(* IEC 61131-3 sources: PLC-ST-Learning/examples/datacenter_control_expert, 5 files *)

(* ---- 01_Types.st ---- *)
(* IEC reference declarations. Create these DDTs in Control Expert's Data Editor.
   This file is NOT an XDB/XEF import file. Indices are always 1..16. *)
TYPE T_DC_TrainStatus :
STRUCT
    Available : BOOL;
    Ready : BOOL;
    Loaded : BOOL;
    ChillerRunning : BOOL;
    Starting : BOOL;
    Stopping : BOOL;
    CanStop : BOOL;
    Fault : BOOL;
    State : INT;
    FaultCode : INT;
END_STRUCT
END_TYPE

TYPE T_DC_StatusArray : ARRAY [1..16] OF T_DC_TrainStatus; END_TYPE
TYPE T_DC_BoolArray : ARRAY [1..16] OF BOOL; END_TYPE
TYPE T_DC_HoursArray : ARRAY [1..16] OF REAL; END_TYPE

TYPE T_DC_TrainIO :
STRUCT
    RemoteAuto : BOOL;
    Maintenance : BOOL;
    RunPermit : BOOL;
    PowerAvailable : BOOL;
    HardTrip : BOOL;
    ChillerFault : BOOL;
    WaterEquipmentFault : BOOL;
    ValveOpenFb : BOOL;
    ValveClosedFb : BOOL;
    ChwPumpRunFb : BOOL;
    CwPumpRunFb : BOOL;
    ChwFlowOk : BOOL;
    CwFlowOk : BOOL;
    TowerReadyFb : BOOL;
    ChillerRunFb : BOOL;
    LoadedFb : BOOL;
    LoadPermit : BOOL;
    Reset : BOOL;
    OpenValvesCmd : BOOL;
    RunChwPumpCmd : BOOL;
    RunCwPumpCmd : BOOL;
    RequestTowerCmd : BOOL;
    RunChillerCmd : BOOL;
    EnableLoadCmd : BOOL;
END_STRUCT
END_TYPE
TYPE T_DC_IOArray : ARRAY [1..16] OF T_DC_TrainIO; END_TYPE

(* ---- 02_FB_DC_Train.st ---- *)
(* Reference DFB: dedicated water equipment per chiller.
   Split declarations and body into a Control Expert DFB; see the Chinese guide.
   All commands are level signals; adapt to vendor start/stop interfaces separately. *)
FUNCTION_BLOCK FB_DC_Train
VAR_INPUT
    FirstScan : BOOL;
    RequestRun : BOOL;
    Reset : BOOL;
    RemoteAuto : BOOL;
    Maintenance : BOOL;
    RunPermit : BOOL;
    PowerAvailable : BOOL; (* Real per-train power feedback, distinct from process trips *)
    HardTrip : BOOL;
    ChillerFault : BOOL;
    WaterEquipmentFault : BOOL;
    ValveOpenFb : BOOL; (* Combined chilled/condenser valve open proof *)
    ValveClosedFb : BOOL;
    ChwPumpRunFb : BOOL;
    CwPumpRunFb : BOOL;
    ChwFlowOk : BOOL;
    CwFlowOk : BOOL;
    TowerReadyFb : BOOL; (* From tower controller; includes local fan staging *)
    ChillerRunFb : BOOL;
    LoadedFb : BOOL; (* Must be real ready/capacity feedback, not command echo *)
    LoadPermit : BOOL;
    MinOff : TIME := T#10m;
    MinOn : TIME := T#10m;
    ValveTimeout : TIME := T#60s;
    PumpTimeout : TIME := T#30s;
    FlowStable : TIME := T#15s;
    FlowTimeout : TIME := T#90s;
    FlowLossDelay : TIME := T#2s;
    CapacityLossDelay : TIME := T#10s;
    TowerTimeout : TIME := T#120s;
    ChillerTimeout : TIME := T#180s;
    LoadTimeout : TIME := T#180s;
    UnloadTimeout : TIME := T#120s;
    StopTimeout : TIME := T#180s;
    PostRun : TIME := T#180s;
END_VAR
VAR_OUTPUT
    OpenValves : BOOL;
    RunChwPump : BOOL;
    RunCwPump : BOOL;
    RequestTower : BOOL;
    RunChiller : BOOL;
    EnableLoad : BOOL;
    Status : T_DC_TrainStatus;
    UnloadTimedOut : BOOL;
    StopTimedOut : BOOL;
END_VAR
VAR
    State : INT;
    FaultLatched : BOOL;
    FaultCode : INT;
    OldReset : BOOL;
    ResetEdge : BOOL;
    WaterOk : BOOL;
    ConfigOk : BOOL;
    ControlledTrip : BOOL;
    tmOff : TON;
    tmOn : TON;
    tmValveOpen : TON;
    tmPump : TON;
    tmFlowStable : TON;
    tmFlowWait : TON;
    tmFlowLoss : TON;
    tmCapacityLoss : TON;
    tmTower : TON;
    tmChiller : TON;
    tmLoad : TON;
    tmUnload : TON;
    tmStop : TON;
    tmPost : TON;
    tmPumpStop : TON;
    tmValveClose : TON;
END_VAR

ResetEdge := Reset AND NOT OldReset;
OldReset := Reset;
ConfigOk := (MinOff > T#0s) AND (MinOn > T#0s)
    AND (ValveTimeout > T#0s) AND (PumpTimeout > T#0s)
    AND (FlowStable > T#0s) AND (FlowTimeout > FlowStable)
    AND (FlowLossDelay >= T#0s) AND (CapacityLossDelay > T#0s)
    AND (TowerTimeout > T#0s)
    AND (ChillerTimeout > T#0s) AND (LoadTimeout > T#0s)
    AND (UnloadTimeout > T#0s) AND (StopTimeout > T#0s)
    AND (PostRun > T#0s);
WaterOk := ValveOpenFb AND ChwPumpRunFb AND CwPumpRunFb
    AND ChwFlowOk AND CwFlowOk;

(* Non-retained state is reconstructed from real feedback, never retained commands. *)
IF FirstScan THEN
    OldReset := Reset;
    ResetEdge := FALSE;
    State := 0;
    FaultLatched := FALSE;
    FaultCode := 0;
    UnloadTimedOut := FALSE;
    StopTimedOut := FALSE;
    IF ChillerRunFb THEN
        IF LoadedFb THEN State := 70; ELSE State := 60; END_IF;
    ELSIF ChwPumpRunFb OR CwPumpRunFb THEN
        State := 100;
    ELSIF ValveOpenFb THEN
        State := 120;
    END_IF;
END_IF;

(* Call EVERY timer exactly once per scan, even while idle or faulted. *)
tmOff(IN := NOT ChillerRunFb AND NOT FirstScan, PT := MinOff);
tmOn(IN := ChillerRunFb AND NOT FirstScan, PT := MinOn);
tmValveOpen(IN := (State = 10) AND NOT FirstScan, PT := ValveTimeout);
tmPump(IN := (State = 20) AND NOT FirstScan, PT := PumpTimeout);
tmFlowStable(IN := WaterOk AND NOT FirstScan, PT := FlowStable);
tmFlowWait(IN := (State = 30) AND NOT FirstScan, PT := FlowTimeout);
tmFlowLoss(IN := (State >= 50) AND (State <= 80) AND NOT WaterOk
    AND NOT FirstScan, PT := FlowLossDelay);
tmCapacityLoss(IN := (State = 70) AND NOT LoadedFb AND NOT FirstScan,
    PT := CapacityLossDelay);
tmTower(IN := (State = 40) AND NOT FirstScan, PT := TowerTimeout);
tmChiller(IN := (State = 50) AND NOT FirstScan, PT := ChillerTimeout);
tmLoad(IN := (State = 60) AND NOT FirstScan, PT := LoadTimeout);
tmUnload(IN := (State = 80) AND NOT FirstScan, PT := UnloadTimeout);
tmStop(IN := (State = 90) AND NOT FirstScan, PT := StopTimeout);
tmPost(IN := (State = 100) AND NOT FirstScan, PT := PostRun);
tmPumpStop(IN := (State = 110) AND NOT FirstScan, PT := PumpTimeout);
tmValveClose(IN := (State = 120) AND NOT FirstScan, PT := ValveTimeout);

IF ResetEdge AND NOT ChillerRunFb AND NOT ChwPumpRunFb AND NOT CwPumpRunFb
    AND ValveClosedFb AND NOT ValveOpenFb AND NOT LoadedFb
    AND NOT ChillerFault AND NOT WaterEquipmentFault AND RunPermit
    AND NOT HardTrip AND RemoteAuto AND PowerAvailable AND ConfigOk
    AND ((State = 0) OR (State = 900)) THEN
    FaultLatched := FALSE;
    FaultCode := 0;
    UnloadTimedOut := FALSE;
    StopTimedOut := FALSE;
    State := 0;
END_IF;

ControlledTrip := FALSE;
IF NOT ConfigOk THEN FaultCode := 1; ControlledTrip := TRUE;
ELSIF NOT RunPermit AND (((State > 0) AND (State < 90)) OR ChillerRunFb) THEN
    FaultCode := 2; ControlledTrip := TRUE;
ELSIF ChillerFault THEN FaultCode := 3; ControlledTrip := TRUE;
ELSIF WaterEquipmentFault THEN FaultCode := 4; ControlledTrip := TRUE;
ELSIF (State >= 50) AND (State <= 80) AND NOT ValveOpenFb THEN
    FaultCode := 5; ControlledTrip := TRUE;
ELSIF tmFlowLoss.Q THEN FaultCode := 6; ControlledTrip := TRUE;
ELSIF (State >= 50) AND (State <= 80) AND NOT TowerReadyFb THEN
    FaultCode := 7; ControlledTrip := TRUE;
ELSIF ((State = 60) OR (State = 70) OR (State = 80)) AND NOT ChillerRunFb THEN
    FaultCode := 8; ControlledTrip := TRUE;
ELSIF tmCapacityLoss.Q THEN
    FaultCode := 9; ControlledTrip := TRUE;
ELSIF LoadedFb AND NOT ChillerRunFb THEN
    FaultCode := 10; ControlledTrip := TRUE;
ELSIF ValveOpenFb AND ValveClosedFb THEN
    FaultCode := 11; ControlledTrip := TRUE;
ELSIF ChillerRunFb AND ((State < 50) OR ((State >= 100) AND (State <= 120))
    OR (State = 900)) THEN
    FaultCode := 14; ControlledTrip := TRUE;
END_IF;

(* Hardwired safeties remain independent. A hard trip removes ALL commands. *)
IF HardTrip THEN
    FaultLatched := TRUE;
    FaultCode := 12;
    State := 900;
ELSIF NOT RemoteAuto THEN
    IF ChillerRunFb OR ChwPumpRunFb OR CwPumpRunFb
        OR ((State > 0) AND (State < 900)) THEN
        FaultLatched := TRUE; FaultCode := 13;
    END_IF;
    IF FaultLatched THEN State := 900; ELSE State := 0; END_IF;
ELSIF NOT PowerAvailable THEN
    (* Expected loss of supply is not a device-fault latch. Existing faults persist. *)
    State := 910;
ELSIF ControlledTrip THEN
    FaultLatched := TRUE;
    IF ChillerRunFb AND (State >= 100) THEN
        State := 90;
    ELSIF (State < 90) OR (State = 900) THEN
        IF ChillerRunFb THEN State := 90;
        ELSIF ChwPumpRunFb OR CwPumpRunFb THEN State := 100;
        ELSIF NOT ValveClosedFb THEN State := 120;
        ELSE State := 900;
        END_IF;
    END_IF;
END_IF;

(* Normal request withdrawal honors MinOn. Startup cancellation needs no MinOn. *)
IF NOT FirstScan AND NOT RequestRun AND NOT ControlledTrip AND NOT HardTrip
    AND RemoteAuto AND PowerAvailable AND (State > 0) AND (State < 80) THEN
    IF (State = 70) AND tmOn.Q THEN State := 80;
    ELSIF State = 10 THEN State := 120;
    ELSIF (State >= 20) AND (State <= 40) THEN State := 100;
    ELSIF (State = 50) OR (State = 60) THEN
        IF ChillerRunFb THEN State := 80; ELSE State := 100; END_IF;
    END_IF;
END_IF;

IF NOT HardTrip AND RemoteAuto AND PowerAvailable THEN
    CASE State OF
    0:
        IF ChillerRunFb OR ChwPumpRunFb OR CwPumpRunFb OR LoadedFb THEN
            FaultLatched := TRUE; FaultCode := 14;
            IF ChillerRunFb THEN State := 90; ELSE State := 100; END_IF;
        ELSIF RequestRun AND NOT FaultLatched AND NOT Maintenance
            AND RunPermit AND ConfigOk AND tmOff.Q AND ValveClosedFb THEN
            State := 10;
        END_IF;
    10:
        IF ValveOpenFb AND NOT ValveClosedFb THEN State := 20;
        ELSIF tmValveOpen.Q THEN FaultLatched := TRUE; FaultCode := 20; State := 120;
        END_IF;
    20:
        IF ChwPumpRunFb AND CwPumpRunFb THEN State := 30;
        ELSIF tmPump.Q THEN FaultLatched := TRUE; FaultCode := 21; State := 100;
        END_IF;
    30:
        IF tmFlowStable.Q THEN State := 40;
        ELSIF tmFlowWait.Q THEN FaultLatched := TRUE; FaultCode := 22; State := 100;
        END_IF;
    40:
        IF TowerReadyFb AND tmFlowStable.Q THEN State := 50;
        ELSIF tmTower.Q THEN FaultLatched := TRUE; FaultCode := 23; State := 100;
        END_IF;
    50:
        IF ChillerRunFb THEN State := 60;
        ELSIF tmChiller.Q THEN FaultLatched := TRUE; FaultCode := 24; State := 90;
        END_IF;
    60:
        IF LoadedFb AND LoadPermit AND tmFlowStable.Q THEN State := 70;
        ELSIF tmLoad.Q THEN FaultLatched := TRUE; FaultCode := 25; State := 80;
        END_IF;
    70:
        (* Loss of load permission unloads through the normal stop path. *)
        IF NOT LoadPermit THEN
            FaultLatched := TRUE; FaultCode := 26; State := 80;
        END_IF;
    80:
        IF NOT LoadedFb THEN State := 90;
        ELSIF tmUnload.Q THEN
            UnloadTimedOut := TRUE; FaultLatched := TRUE; FaultCode := 27; State := 90;
        END_IF;
    90:
        (* A stuck run feedback MUST NOT be treated as a stopped chiller. *)
        IF NOT ChillerRunFb THEN State := 100;
        ELSIF tmStop.Q THEN
            StopTimedOut := TRUE; FaultLatched := TRUE; FaultCode := 28;
        END_IF;
    100:
        IF ChillerRunFb THEN
            FaultLatched := TRUE; FaultCode := 29; State := 90;
        ELSIF tmPost.Q THEN State := 110;
        END_IF;
    110:
        IF NOT ChwPumpRunFb AND NOT CwPumpRunFb THEN State := 120;
        ELSIF tmPumpStop.Q THEN
            FaultLatched := TRUE; FaultCode := 30;
            (* Keep valves open until BOTH pumps really stop. *)
        END_IF;
    120:
        IF ChillerRunFb OR ChwPumpRunFb OR CwPumpRunFb THEN
            FaultLatched := TRUE; FaultCode := 31;
            IF ChillerRunFb THEN State := 90; ELSE State := 110; END_IF;
        ELSIF ValveClosedFb AND NOT ValveOpenFb THEN
            IF FaultLatched THEN State := 900; ELSE State := 0; END_IF;
        ELSIF tmValveClose.Q THEN
            FaultLatched := TRUE; FaultCode := 32;
        END_IF;
    900:
        (* No automatic reset/retry. A real reset edge at a safe rest is required. *)
        IF ChillerRunFb THEN State := 90;
        ELSIF ChwPumpRunFb OR CwPumpRunFb THEN State := 100;
        END_IF;
    910:
        (* Re-establish a safe rest before allowing the fleet to restart this train. *)
        IF ChillerRunFb THEN State := 90;
        ELSIF ChwPumpRunFb OR CwPumpRunFb THEN State := 100;
        ELSIF NOT ValveClosedFb THEN State := 120;
        ELSIF FaultLatched THEN State := 900;
        ELSE State := 0;
        END_IF;
    ELSE
        FaultLatched := TRUE; FaultCode := 99;
        IF ChillerRunFb THEN State := 90; ELSE State := 100; END_IF;
    END_CASE;
END_IF;

OpenValves := (State >= 10) AND (State <= 110);
RunChwPump := (State >= 20) AND (State <= 100);
RunCwPump := RunChwPump;
RequestTower := (State >= 40) AND (State <= 100);
RunChiller := (State >= 50) AND (State <= 80);
EnableLoad := (((State = 60) AND tmFlowStable.Q) OR ((State = 70) AND WaterOk))
    AND LoadPermit AND TowerReadyFb AND ChillerRunFb AND NOT FaultLatched;
(* Physical interlocks cut chiller/load immediately; water may continue for post-run. *)
RunChiller := RunChiller AND RunPermit AND NOT ChillerFault
    AND NOT WaterEquipmentFault AND ValveOpenFb AND NOT tmFlowLoss.Q
    AND TowerReadyFb AND ConfigOk AND ((State <> 50) OR WaterOk);
IF HardTrip OR NOT RemoteAuto OR NOT PowerAvailable THEN
    OpenValves := FALSE; RunChwPump := FALSE; RunCwPump := FALSE;
    RequestTower := FALSE; RunChiller := FALSE; EnableLoad := FALSE;
END_IF;
EnableLoad := EnableLoad AND RunChiller;
Status.Available := RemoteAuto AND NOT Maintenance AND RunPermit
    AND PowerAvailable
    AND NOT HardTrip AND NOT ChillerFault AND NOT WaterEquipmentFault
    AND NOT FaultLatched AND ConfigOk;
Status.Ready := Status.Available AND (State = 0) AND tmOff.Q
    AND ValveClosedFb AND NOT ValveOpenFb AND NOT ChillerRunFb
    AND NOT ChwPumpRunFb AND NOT CwPumpRunFb AND NOT LoadedFb;
Status.Loaded := (State = 70) AND LoadedFb AND ChillerRunFb AND WaterOk
    AND TowerReadyFb AND LoadPermit AND NOT FaultLatched
    AND RemoteAuto AND RunPermit AND NOT HardTrip;
Status.ChillerRunning := ChillerRunFb;
Status.Starting := (State >= 10) AND (State <= 60);
Status.Stopping := (State >= 80) AND (State <= 120);
Status.CanStop := (State = 70) AND tmOn.Q;
Status.Fault := FaultLatched;
Status.State := State;
Status.FaultCode := FaultCode;
END_FUNCTION_BLOCK

(* ---- 03_FB_DC_Plant.st ---- *)
(* Fleet dispatch. Equal-capacity chillers; maximum 16.
   Call all Train DFBs BEFORE this DFB; requests take effect next PLC scan. *)
FUNCTION_BLOCK FB_DC_Plant
VAR_INPUT
    FirstScan : BOOL;
    Enable : BOOL;
    DisasterActive : BOOL; (* Recovery latch input, NOT a safety output *)
    InfrastructureReady : BOOL; (* Power, BMS authority, common water system ready *)
    AckRecovery : BOOL;
    AutoRecovery : BOOL := FALSE;
    ResetAlarm : BOOL;
    DemandValid : BOOL;
    Demand : INT; (* Desired duty count from BMS or validated demand regulator *)
    UnitCount : INT := 4;
    MaxDuty : INT := 3; (* N+1 reserve with four installed units *)
    MaxParallel : INT := 4; (* Electrical/hydraulic limit, includes rotation overlap *)
    RotateEnable : BOOL := TRUE;
    RotateNow : BOOL;
    Status : T_DC_StatusArray;
    RunHours : T_DC_HoursArray; (* External, validated RETAIN hour meters *)
    RecoveryStable : TIME := T#60s;
    StartSpacing : TIME := T#120s;
    DemandUpDelay : TIME := T#60s;
    DemandDownDelay : TIME := T#300s;
    RotationInterval : TIME := T#168h;
    RotationOverlap : TIME := T#60s;
    RotationTimeout : TIME := T#30m;
END_VAR
VAR_OUTPUT
    Request : T_DC_BoolArray;
    RecoveryHold : BOOL;
    Target : INT;
    RunningCount : INT;
    LoadedCount : INT;
    RequestedCount : INT;
    CapacityShortage : BOOL;
    NoStartCandidate : BOOL;
    ReserveUnavailable : BOOL;
    ConfigFault : BOOL;
    RotationBlocked : BOOL;
    RotationFailed : BOOL;
    RotationActive : BOOL;
    InvalidDemand : BOOL;
END_VAR
VAR
    i : INT;
    n : INT;
    Candidate : INT;
    StopCandidate : INT;
    RotOld : INT;
    RotNew : INT;
    RotPhase : INT; (* 0 idle; 1 start replacement; 2 old train shutting down *)
    ReadyCount : INT;
    OccupiedCount : INT;
    LastDemand : INT;
    RotationTarget : INT;
    Desired : INT;
    MinHours : REAL;
    MaxHours : REAL;
    Starting : BOOL;
    Stopping : BOOL;
    OldAck : BOOL;
    OldRotate : BOOL;
    OldReset : BOOL;
    AckEdge : BOOL;
    RotateEdge : BOOL;
    ResetEdge : BOOL;
    SpacingActive : BOOL;
    SpacingReset : BOOL;
    RotationClockReset : BOOL;
    ReplacementLoaded : BOOL;
    tmRecovery : TON;
    tmSpacing : TON;
    tmUp : TON;
    tmDown : TON;
    tmRotation : TON;
    tmOverlap : TON;
    tmRotationTimeout : TON;
END_VAR

ConfigFault := (UnitCount < 1) OR (UnitCount > 16) OR (MaxDuty < 1)
    OR (MaxDuty > UnitCount) OR (MaxParallel < MaxDuty)
    OR (MaxParallel > UnitCount) OR (RecoveryStable <= T#0s)
    OR (StartSpacing <= T#0s) OR (DemandUpDelay < T#0s)
    OR (DemandDownDelay < T#0s) OR (RotationInterval <= T#0s)
    OR (RotationOverlap <= T#0s) OR (RotationTimeout <= RotationOverlap);
n := UnitCount;
IF n < 1 THEN n := 1; END_IF;
IF n > 16 THEN n := 16; END_IF;
AckEdge := AckRecovery AND NOT OldAck;
RotateEdge := RotateNow AND NOT OldRotate;
ResetEdge := ResetAlarm AND NOT OldReset;
OldAck := AckRecovery; OldRotate := RotateNow; OldReset := ResetAlarm;

IF FirstScan THEN
    RecoveryHold := TRUE;
    Target := 0; LastDemand := -1;
    RotPhase := 0; RotOld := 0; RotNew := 0;
    SpacingActive := TRUE; SpacingReset := TRUE; RotationClockReset := TRUE;
    RotationFailed := FALSE;
    AckEdge := FALSE; RotateEdge := FALSE; ResetEdge := FALSE;
    (* Adopt operating trains; never replay a retained command array. *)
    FOR i := 1 TO 16 DO
        Request[i] := (i <= n) AND Status[i].Available
            AND (Status[i].ChillerRunning OR Status[i].Starting);
        IF Request[i] THEN Target := Target + 1; END_IF;
    END_FOR;
END_IF;
IF DisasterActive OR NOT InfrastructureReady THEN RecoveryHold := TRUE; END_IF;

(* Invalid demand freezes the current target; it MUST NOT become zero demand. *)
InvalidDemand := NOT DemandValid OR (Demand < 0) OR (Demand > MaxDuty);
Desired := Target;
IF NOT InvalidDemand THEN Desired := Demand; END_IF;
IF NOT Enable THEN Desired := 0; END_IF;

tmRecovery(IN := InfrastructureReady AND NOT DisasterActive AND NOT FirstScan,
    PT := RecoveryStable);
tmSpacing(IN := SpacingActive AND NOT SpacingReset AND NOT FirstScan, PT := StartSpacing);
tmUp(IN := Enable AND NOT InvalidDemand AND NOT RecoveryHold
    AND (Desired > Target) AND (Desired = LastDemand) AND NOT FirstScan,
    PT := DemandUpDelay);
tmDown(IN := NOT InvalidDemand AND NOT RecoveryHold AND (Desired < Target)
    AND (Desired = LastDemand) AND NOT FirstScan, PT := DemandDownDelay);
tmRotation(IN := Enable AND RotateEnable AND NOT RecoveryHold AND (Target > 0)
    AND (RotPhase = 0) AND NOT RotationClockReset AND NOT FirstScan,
    PT := RotationInterval);
ReplacementLoaded := FALSE;
IF (RotNew >= 1) AND (RotNew <= n) THEN
    ReplacementLoaded := Status[RotNew].Loaded;
END_IF;
tmOverlap(IN := (RotPhase = 1) AND ReplacementLoaded
    AND NOT FirstScan, PT := RotationOverlap);
tmRotationTimeout(IN := (RotPhase <> 0) AND NOT FirstScan, PT := RotationTimeout);
RotationClockReset := FALSE;
SpacingReset := FALSE;
IF tmSpacing.Q THEN SpacingActive := FALSE; END_IF;
IF ResetEdge THEN RotationFailed := FALSE; END_IF;
IF RecoveryHold AND tmRecovery.Q AND (AutoRecovery OR AckEdge) AND Enable
    AND NOT ConfigFault THEN
    RecoveryHold := FALSE;
    SpacingActive := TRUE;
    SpacingReset := TRUE;
END_IF;
IF NOT Enable THEN Target := 0;
ELSIF NOT RecoveryHold AND NOT ConfigFault THEN
    IF tmUp.Q OR tmDown.Q THEN Target := Desired; END_IF;
END_IF;
LastDemand := Desired;

RunningCount := 0; LoadedCount := 0; RequestedCount := 0;
ReadyCount := 0; OccupiedCount := 0;
Starting := FALSE; Stopping := FALSE;
FOR i := 1 TO 16 DO
    IF i <= n THEN
        IF Status[i].ChillerRunning THEN RunningCount := RunningCount + 1; END_IF;
        IF Status[i].Loaded THEN LoadedCount := LoadedCount + 1; END_IF;
        IF Status[i].Ready THEN ReadyCount := ReadyCount + 1; END_IF;
        IF NOT Status[i].Available THEN Request[i] := FALSE; END_IF;
        IF Request[i] THEN RequestedCount := RequestedCount + 1; END_IF;
        IF Request[i] OR Status[i].ChillerRunning OR Status[i].Starting THEN
            OccupiedCount := OccupiedCount + 1;
        END_IF;
        Starting := Starting OR Status[i].Starting;
        Stopping := Stopping OR Status[i].Stopping;
    ELSE
        Request[i] := FALSE;
    END_IF;
END_FOR;

(* Select least-hours available start and greatest-hours stoppable running train.
   Ascending index resolves ties deterministically. *)
Candidate := 0; StopCandidate := 0;
MinHours := 3.0E+38; MaxHours := -1.0;
FOR i := 1 TO n DO
    IF Status[i].Ready AND NOT Request[i] AND (RunHours[i] >= 0.0)
        AND (RunHours[i] < MinHours) THEN
        Candidate := i; MinHours := RunHours[i];
    END_IF;
    IF Request[i] AND Status[i].Loaded AND Status[i].CanStop
        AND (RunHours[i] >= 0.0) AND (RunHours[i] > MaxHours) THEN
        StopCandidate := i; MaxHours := RunHours[i];
    END_IF;
END_FOR;

RotationBlocked := FALSE;
IF RotPhase <> 0 THEN
    (* Bound indices before use. No reliance on short-circuit array evaluation. *)
    IF (RotOld < 1) OR (RotOld > n) OR (RotNew < 1) OR (RotNew > n) THEN
        RotPhase := 0; RotationFailed := TRUE; RotationClockReset := TRUE;
    ELSE
        IF ConfigFault OR RecoveryHold OR NOT Enable OR InvalidDemand
            OR (Target <> RotationTarget) THEN
            (* Keep the original running unit; cancel replacement normally. *)
            IF RotPhase = 1 THEN Request[RotNew] := FALSE; END_IF;
            RotPhase := 0; RotationClockReset := TRUE;
        ELSIF NOT Status[RotOld].Available THEN
            (* Original failed: replacement is now ordinary fault replacement. *)
            RotPhase := 0; RotationClockReset := TRUE;
        ELSIF NOT Status[RotNew].Available OR tmRotationTimeout.Q THEN
            IF RotPhase = 1 THEN Request[RotNew] := FALSE; END_IF;
            RotationFailed := TRUE; RotPhase := 0; RotationClockReset := TRUE;
        ELSIF RotPhase = 1 THEN
            IF Status[RotNew].Loaded AND tmOverlap.Q AND Status[RotOld].CanStop THEN
                Request[RotOld] := FALSE; RotPhase := 2;
            END_IF;
        ELSIF RotPhase = 2 THEN
            IF NOT Status[RotOld].ChillerRunning AND NOT Status[RotOld].Stopping THEN
                RotPhase := 0; RotationClockReset := TRUE;
            END_IF;
        END_IF;
    END_IF;
END_IF;

IF NOT ConfigFault AND NOT RecoveryHold AND Enable
    AND (RotPhase = 0) AND NOT Starting THEN
    IF RequestedCount < Target THEN
        (* Fault replacement bypasses demand debounce, not start spacing or MinOff.
           Failed trains may finish water post-run while a spare starts. *)
        IF (Candidate > 0) AND NOT SpacingActive AND (OccupiedCount < MaxParallel) THEN
            Request[Candidate] := TRUE;
            SpacingActive := TRUE;
            SpacingReset := TRUE;
        END_IF;
    ELSIF (RequestedCount > Target) AND NOT Stopping AND NOT InvalidDemand THEN
        IF StopCandidate > 0 THEN Request[StopCandidate] := FALSE; END_IF;
    ELSIF RotateEnable AND NOT InvalidDemand AND (RotateEdge OR tmRotation.Q) AND (Target > 0)
        AND (RequestedCount = Target) AND (LoadedCount >= Target)
        AND NOT Stopping THEN
        IF (Candidate > 0) AND (StopCandidate > 0) AND NOT SpacingActive
            AND (OccupiedCount < MaxParallel) THEN
            RotOld := StopCandidate; RotNew := Candidate; RotationTarget := Target;
            Request[RotNew] := TRUE; RotPhase := 1; SpacingActive := TRUE;
            SpacingReset := TRUE;
            RotationClockReset := TRUE;
        ELSE RotationBlocked := TRUE;
        END_IF;
    END_IF;
END_IF;
(* Disable is an orderly stop; hard stops are the individual Train.HardTrip input. *)
IF NOT Enable THEN
    FOR i := 1 TO 16 DO Request[i] := FALSE; END_FOR;
END_IF;

RotationActive := RotPhase <> 0;
RequestedCount := 0;
FOR i := 1 TO n DO
    IF Request[i] THEN RequestedCount := RequestedCount + 1; END_IF;
END_FOR;
CapacityShortage := Enable AND NOT InvalidDemand AND (LoadedCount < Demand);
NoStartCandidate := Enable AND NOT RecoveryHold
    AND (RequestedCount < Target) AND (Candidate = 0);
ReserveUnavailable := Enable AND (ReadyCount = 0);
END_FUNCTION_BLOCK

(* ---- 04_FB_DC_Demand.st ---- *)
(* Optional supervisory staging by chilled-water SUPPLY temperature.
   Native chiller controllers retain compressor/guide-vane/VFD modulation.
   Do not use with unequal-capacity units without a capacity-based redesign. *)
FUNCTION_BLOCK FB_DC_Demand
VAR_INPUT
    FirstScan : BOOL;
    Enable : BOOL;
    SensorValid : BOOL;
    SupplyTemperature : REAL;
    Setpoint : REAL := 7.0;
    AddBand : REAL := 0.7;
    ShedBand : REAL := 0.5;
    SensorMin : REAL := 0.0;
    SensorMax : REAL := 35.0;
    MinDuty : INT := 1;
    MaxDuty : INT := 3;
    LoadedCount : INT;
    PlantStable : BOOL; (* No starts, stops, rotation, or recovery in progress *)
    AddDelay : TIME := T#120s;
    ShedDelay : TIME := T#600s;
    SettleTime : TIME := T#600s;
END_VAR
VAR_OUTPUT
    Demand : INT;
    DemandValid : BOOL;
    SensorAlarm : BOOL;
    ConfigFault : BOOL;
END_VAR
VAR
    tmAdd : TON;
    tmShed : TON;
    tmSettle : TON;
    Settling : BOOL;
    ResetSettle : BOOL;
    CanAdjust : BOOL;
END_VAR

ConfigFault := (MinDuty < 0) OR (MaxDuty < 1) OR (MaxDuty > 16)
    OR (MinDuty > MaxDuty) OR (AddBand <= 0.0) OR (ShedBand <= 0.0)
    OR (SensorMin >= SensorMax) OR (Setpoint <= SensorMin)
    OR (Setpoint >= SensorMax) OR (AddDelay <= T#0s)
    OR (ShedDelay <= T#0s) OR (SettleTime <= T#0s);
(* Positive range tests also reject an IEEE NaN measurement. *)
SensorAlarm := NOT SensorValid OR NOT ((SupplyTemperature >= SensorMin)
    AND (SupplyTemperature <= SensorMax));
DemandValid := NOT ConfigFault AND NOT SensorAlarm;
IF FirstScan THEN
    Demand := MinDuty;
    IF (LoadedCount > MinDuty) AND (LoadedCount <= MaxDuty) THEN
        Demand := LoadedCount;
    END_IF;
    IF Demand < 0 THEN Demand := 0; END_IF;
    IF Demand > 16 THEN Demand := 16; END_IF;
    Settling := TRUE; ResetSettle := TRUE;
END_IF;
tmSettle(IN := Settling AND NOT ResetSettle AND NOT FirstScan, PT := SettleTime);
ResetSettle := FALSE;
IF tmSettle.Q THEN Settling := FALSE; END_IF;
CanAdjust := Enable AND DemandValid AND PlantStable AND NOT Settling
    AND (LoadedCount = Demand) AND NOT FirstScan;
tmAdd(IN := CanAdjust AND (SupplyTemperature > Setpoint + AddBand)
    AND (Demand < MaxDuty), PT := AddDelay);
tmShed(IN := CanAdjust AND (SupplyTemperature < Setpoint - ShedBand)
    AND (Demand > MinDuty), PT := ShedDelay);
IF NOT Enable THEN
    Demand := 0; Settling := TRUE; ResetSettle := TRUE;
ELSIF DemandValid THEN
    IF Demand < MinDuty THEN
        Demand := MinDuty; Settling := TRUE; ResetSettle := TRUE;
    ELSIF Demand > MaxDuty THEN
        Demand := MaxDuty; Settling := TRUE; ResetSettle := TRUE;
    ELSIF tmAdd.Q THEN
        Demand := Demand + 1; Settling := TRUE; ResetSettle := TRUE;
    ELSIF tmShed.Q THEN
        Demand := Demand - 1; Settling := TRUE; ResetSettle := TRUE;
    END_IF;
END_IF;
(* With invalid measurement Demand is held, not forced to zero. *)
END_FUNCTION_BLOCK

(* ---- 05_PRG_DC_Example.st ---- *)
(* Four equal-capacity water-cooled chillers, each with dedicated pumps/valves.
   REFERENCE ONLY: create DDTs, DFBs and application variables in Control Expert.
   Split PROGRAM declarations/body into Data Editor + periodic MAST ST section.
   Map IO from/to field adapters BEFORE/AFTER this section respectively.
   ColdOrWarmStart must pulse for every PLC restart; see guide. *)
PROGRAM PRG_DC_Example
VAR
    ColdOrWarmStart : BOOL;
    FirstScan : BOOL;
    InitDone : BOOL;
    AutoEnable : BOOL;
    DisasterActive : BOOL;
    InfrastructureReady : BOOL;
    RecoveryAcknowledgement : BOOL;
    AlarmReset : BOOL;
    RotateCommand : BOOL;
    TemperatureQualityGood : BOOL;
    SupplyTemperature : REAL;
    IO : T_DC_IOArray;
    UnitStatus : T_DC_StatusArray;
    RunHours : T_DC_HoursArray;
    Requests : T_DC_BoolArray;
    Train01 : FB_DC_Train;
    Train02 : FB_DC_Train;
    Train03 : FB_DC_Train;
    Train04 : FB_DC_Train;
    Plant : FB_DC_Plant;
    DemandRegulator : FB_DC_Demand;
    ActualLoaded : INT;
    PlantStable : BOOL;
    i : INT;
END_VAR

FirstScan := ColdOrWarmStart OR NOT InitDone;
InitDone := TRUE;

Train01(FirstScan := FirstScan, RequestRun := Requests[1],
    RemoteAuto := IO[1].RemoteAuto,
    Maintenance := IO[1].Maintenance,
    RunPermit := IO[1].RunPermit,
    PowerAvailable := IO[1].PowerAvailable,
    HardTrip := IO[1].HardTrip,
    ChillerFault := IO[1].ChillerFault,
    WaterEquipmentFault := IO[1].WaterEquipmentFault,
    ValveOpenFb := IO[1].ValveOpenFb,
    ValveClosedFb := IO[1].ValveClosedFb,
    ChwPumpRunFb := IO[1].ChwPumpRunFb,
    CwPumpRunFb := IO[1].CwPumpRunFb,
    ChwFlowOk := IO[1].ChwFlowOk,
    CwFlowOk := IO[1].CwFlowOk,
    TowerReadyFb := IO[1].TowerReadyFb,
    ChillerRunFb := IO[1].ChillerRunFb,
    LoadedFb := IO[1].LoadedFb,
    LoadPermit := IO[1].LoadPermit,
    Reset := IO[1].Reset);
IO[1].OpenValvesCmd := Train01.OpenValves;
IO[1].RunChwPumpCmd := Train01.RunChwPump;
IO[1].RunCwPumpCmd := Train01.RunCwPump;
IO[1].RequestTowerCmd := Train01.RequestTower;
IO[1].RunChillerCmd := Train01.RunChiller;
IO[1].EnableLoadCmd := Train01.EnableLoad;
UnitStatus[1] := Train01.Status;

Train02(FirstScan := FirstScan, RequestRun := Requests[2],
    RemoteAuto := IO[2].RemoteAuto,
    Maintenance := IO[2].Maintenance,
    RunPermit := IO[2].RunPermit,
    PowerAvailable := IO[2].PowerAvailable,
    HardTrip := IO[2].HardTrip,
    ChillerFault := IO[2].ChillerFault,
    WaterEquipmentFault := IO[2].WaterEquipmentFault,
    ValveOpenFb := IO[2].ValveOpenFb,
    ValveClosedFb := IO[2].ValveClosedFb,
    ChwPumpRunFb := IO[2].ChwPumpRunFb,
    CwPumpRunFb := IO[2].CwPumpRunFb,
    ChwFlowOk := IO[2].ChwFlowOk,
    CwFlowOk := IO[2].CwFlowOk,
    TowerReadyFb := IO[2].TowerReadyFb,
    ChillerRunFb := IO[2].ChillerRunFb,
    LoadedFb := IO[2].LoadedFb,
    LoadPermit := IO[2].LoadPermit,
    Reset := IO[2].Reset);
IO[2].OpenValvesCmd := Train02.OpenValves;
IO[2].RunChwPumpCmd := Train02.RunChwPump;
IO[2].RunCwPumpCmd := Train02.RunCwPump;
IO[2].RequestTowerCmd := Train02.RequestTower;
IO[2].RunChillerCmd := Train02.RunChiller;
IO[2].EnableLoadCmd := Train02.EnableLoad;
UnitStatus[2] := Train02.Status;

Train03(FirstScan := FirstScan, RequestRun := Requests[3],
    RemoteAuto := IO[3].RemoteAuto,
    Maintenance := IO[3].Maintenance,
    RunPermit := IO[3].RunPermit,
    PowerAvailable := IO[3].PowerAvailable,
    HardTrip := IO[3].HardTrip,
    ChillerFault := IO[3].ChillerFault,
    WaterEquipmentFault := IO[3].WaterEquipmentFault,
    ValveOpenFb := IO[3].ValveOpenFb,
    ValveClosedFb := IO[3].ValveClosedFb,
    ChwPumpRunFb := IO[3].ChwPumpRunFb,
    CwPumpRunFb := IO[3].CwPumpRunFb,
    ChwFlowOk := IO[3].ChwFlowOk,
    CwFlowOk := IO[3].CwFlowOk,
    TowerReadyFb := IO[3].TowerReadyFb,
    ChillerRunFb := IO[3].ChillerRunFb,
    LoadedFb := IO[3].LoadedFb,
    LoadPermit := IO[3].LoadPermit,
    Reset := IO[3].Reset);
IO[3].OpenValvesCmd := Train03.OpenValves;
IO[3].RunChwPumpCmd := Train03.RunChwPump;
IO[3].RunCwPumpCmd := Train03.RunCwPump;
IO[3].RequestTowerCmd := Train03.RequestTower;
IO[3].RunChillerCmd := Train03.RunChiller;
IO[3].EnableLoadCmd := Train03.EnableLoad;
UnitStatus[3] := Train03.Status;

Train04(FirstScan := FirstScan, RequestRun := Requests[4],
    RemoteAuto := IO[4].RemoteAuto,
    Maintenance := IO[4].Maintenance,
    RunPermit := IO[4].RunPermit,
    PowerAvailable := IO[4].PowerAvailable,
    HardTrip := IO[4].HardTrip,
    ChillerFault := IO[4].ChillerFault,
    WaterEquipmentFault := IO[4].WaterEquipmentFault,
    ValveOpenFb := IO[4].ValveOpenFb,
    ValveClosedFb := IO[4].ValveClosedFb,
    ChwPumpRunFb := IO[4].ChwPumpRunFb,
    CwPumpRunFb := IO[4].CwPumpRunFb,
    ChwFlowOk := IO[4].ChwFlowOk,
    CwFlowOk := IO[4].CwFlowOk,
    TowerReadyFb := IO[4].TowerReadyFb,
    ChillerRunFb := IO[4].ChillerRunFb,
    LoadedFb := IO[4].LoadedFb,
    LoadPermit := IO[4].LoadPermit,
    Reset := IO[4].Reset);
IO[4].OpenValvesCmd := Train04.OpenValves;
IO[4].RunChwPumpCmd := Train04.RunChwPump;
IO[4].RunCwPumpCmd := Train04.RunCwPump;
IO[4].RequestTowerCmd := Train04.RequestTower;
IO[4].RunChillerCmd := Train04.RunChiller;
IO[4].EnableLoadCmd := Train04.EnableLoad;
UnitStatus[4] := Train04.Status;

ActualLoaded := 0;
PlantStable := NOT Plant.RecoveryHold AND NOT Plant.RotationActive;
FOR i := 1 TO 4 DO
    IF UnitStatus[i].Loaded THEN ActualLoaded := ActualLoaded + 1; END_IF;
    PlantStable := PlantStable AND NOT UnitStatus[i].Starting AND NOT UnitStatus[i].Stopping;
END_FOR;

DemandRegulator(
    FirstScan := FirstScan, Enable := AutoEnable,
    SensorValid := TemperatureQualityGood, SupplyTemperature := SupplyTemperature,
    LoadedCount := ActualLoaded, PlantStable := PlantStable,
    MinDuty := 1, MaxDuty := 3);

Plant(
    FirstScan := FirstScan, Enable := AutoEnable,
    DisasterActive := DisasterActive, InfrastructureReady := InfrastructureReady,
    AckRecovery := RecoveryAcknowledgement, AutoRecovery := FALSE,
    ResetAlarm := AlarmReset, DemandValid := DemandRegulator.DemandValid,
    Demand := DemandRegulator.Demand, UnitCount := 4, MaxDuty := 3, MaxParallel := 4,
    RotateEnable := TRUE, RotateNow := RotateCommand,
    Status := UnitStatus, RunHours := RunHours);
Requests := Plant.Request;

(* HMI: expose all UnitStatus fields, Plant outputs, Train unload/stop timeout
   alarms, and DemandRegulator.SensorAlarm / ConfigFault.
   IO is a software image: physical output writing and vendor protocol adapters
   belong to the application's single-authority I/O layer. *)
END_PROGRAM
